(* IEC 61131-3 sources: programs/VI-54/VI-54_20171205/VI-54_20171205/Stations/PLC_VI54/VI-54_171014/Class/_DriveASyncPara, 1 file *)

(* ---- _DriveASyncPara.st ---- *)
#include "..\..\Class\_DriveMngBase\SDDDefinitions.h"

(*!
<Class
	Name               = "_DriveASyncPara"
	Revision           = "1.2"
	RealtimeTask       = "false"
	CyclicTask         = "false"
	BackgroundTask     = "false"
	Sigmatek           = "true"
	OSInterface        = "false"
	HighPriority       = "false"
	Automatic          = "false"
	UpdateMode         = "Prescan"
	IconPath           = ".\Class\_DriveMngBase\Drive.ico"
	SharedCommandTable = "true"
	Objectsize         = "(330,120)"
	Comment            = "class for asynchron parameter handling">
	<Channels>
		<Server Name="ErrorQuit" Visualized="true" Initialize="false" WriteProtected="false" Retentive="false" Comment="quit an error if the asnychron parameter handling failed"/>
		<Server Name="ParaNr" Visualized="true" Initialize="false" WriteProtected="false" Retentive="false" Comment="write the parameter number to read/write the value"/>
		<Server Name="ParaRdWr" Visualized="true" Initialize="false" WriteProtected="false" Retentive="false" Comment="0 .. read the value of the parameter number&#13;&#10;1 .. write a new value of the parameter number"/>
		<Server Name="ParaValue" Visualized="true" Initialize="false" WriteProtected="false" Retentive="false" Comment="Read Command = actual value of the parameter&#13;&#10;Write Command = the new value which has to written to the parameter"/>
		<Server Name="State" Visualized="true" Initialize="false" WriteProtected="true" Retentive="false" Comment="Actual state of the asynchron handling class&#13;&#10;Following states are possible :&#13;&#10;READY&#13;&#10;BUSY&#13;&#10;ERROR"/>
		<Client Name="DriveAxis" Required="true" Internal="false" Comment="object channel to the class _DriveAxis"/>
		<Client Name="ErrorCode" Required="false" Internal="false" Comment="Following error codes are possible :&#13;&#10;ErrorCode &#13;&#10;   3 =    object change only in disable state&#13;&#10;   4 =    object value greater max value or smaller min value&#13;&#10;   5 =    object write not possible&#13;&#10;   6 =    object cannot be changed in this mode&#13;&#10;   7 =    object not available&#13;&#10;   8 =    object read not possible&#13;&#10;   9 =    initialisation processed successful&#13;&#10;  10 =    communication not initialised&#13;&#10;  11 =    axis is not available&#13;&#10;&#13;&#10;"/>
	</Channels>
	<Dependencies>
		<Files>
			<File Path=".\Class\_DriveMngBase\SDDDefinitions.h" Include="true"/>
		</Files>
	</Dependencies>
	<RevDoku>
		<Owner Company="Sigmatek" Author="HasHan"/>
		<Dokumentation Revision="1.2" Date="17.09.2012" Author="RamAnd" Company="Sigmatek" Description="Added method IsOnline to check online state before starting a request."/>
		<Dokumentation Revision="1.1" Date="21.07.2011" Author="RamAnd" Company="Sigmatek" Description="Changed object client DriveAxis from class _DriveAxis to _DriveAxisBase, like in all other drive classes with a connection to the axis object."/>
		<Dokumentation Revision="1.0" Date="05.08.2009" Author="HasHan" Company="Sigmatek" Description="Creation"/>
	</RevDoku>
</Class>
*)
_DriveASyncPara : CLASS
  //Servers:
	State 	: SvrChCmd_iprStates;
	ParaNr 	: SvrCh_DINT;
	ParaRdWr 	: SvrCh_DINT;
	ParaValue 	: SvrCh_DINT;
	ErrorQuit 	: SvrCh_DINT;
  //Clients:
	DriveAxis 	: CltChCmd__DriveAxisBase;
	ErrorCode 	: CltCh_DINT;
  //Variables:
  //Functions:

	FUNCTION VIRTUAL GLOBAL Init;
				//! <Function Comment="get the online state (checks if the axis module can be accessed)" Name="IsOnline"/>
	FUNCTION GLOBAL IsOnline
		VAR_OUTPUT
			OnlineState 	: DINT;			//! <Variable Comment="0..offline&#13;&#10;1..online" Name="IsOnline.OnlineState"/>
		END_VAR;

	FUNCTION VIRTUAL GLOBAL State::NewInst
		VAR_INPUT
			pPara 	: ^CmdStruct;
			pResult 	: ^results;
		END_VAR
		VAR_OUTPUT
			ret_code 	: iprStates;
		END_VAR;

	FUNCTION VIRTUAL GLOBAL ParaNr::Write
		VAR_INPUT
			input (EAX) 	: DINT;
		END_VAR
		VAR_OUTPUT
			result (EAX) 	: DINT;
		END_VAR;

	FUNCTION VIRTUAL GLOBAL ErrorQuit::Write
		VAR_INPUT
			input (EAX) 	: DINT;
		END_VAR
		VAR_OUTPUT
			result (EAX) 	: DINT;
		END_VAR;
  //Tables:
	FUNCTION @STD
		VAR_OUTPUT
			ret_code	: CONFSTATES;
		END_VAR;
	FUNCTION GLOBAL TAB @CT_;
END_CLASS;

#pragma usingLtd _DriveAxisBase

FUNCTION VIRTUAL GLOBAL _DriveASyncPara::Init

	if _firstscan then
    State := READY;
    ErrorCode := 0;
	end_if;

END_FUNCTION

FUNCTION VIRTUAL GLOBAL _DriveASyncPara::State::NewInst
	VAR_INPUT
		pPara 	: ^CmdStruct;
		pResult 	: ^results;
	END_VAR
	VAR_OUTPUT
		ret_code 	: iprStates;
	END_VAR

	ret_code:= READY;

	case pPara^.uiCmd of
	SDD_ASYNC_READY :
		// was the command a read or a write command
		if pPara^.aPara[1] = 0 then
			// read command
			ParaValue := pPara^.aPara[2];
		end_if;
		State := READY;

  SDD_ASYNC_ERROR :
    ErrorCode := pPara^.aPara[1];
    ErrorCode.write(ErrorCode);
    State := ERROR;

	end_case;

END_FUNCTION

FUNCTION VIRTUAL GLOBAL _DriveASyncPara::ParaNr::Write
	VAR_INPUT
		input (EAX) 	: DINT;
	END_VAR
	VAR_OUTPUT
		result (EAX) 	: DINT;
	END_VAR
  VAR
  	IntState    : iprStates;
  END_VAR

	result := ACCESS_DENIED;

	if (State = READY) then
		ParaNr := input;
    IntState := DriveAxis.CmdState.Read();

    if IntState = ERROR then
      if DriveAxis.AxisState.NoHW = 1 then
        ErrorCode := 11;
        ErrorCode.write(ErrorCode);
      end_if;
      State := DriveAxis := IntState;
      return;
    end_if;

		// Add the entry into the ring buffer
		result := DriveAxis.AddASyncEntry(to_usint(ParaNr), to_usint(ParaRdWr), ParaValue, this, 0);
		if result = 0 then
			State := BUSY;
		end_if;
	end_if;

END_FUNCTION

FUNCTION VIRTUAL GLOBAL _DriveASyncPara::ErrorQuit::Write
	VAR_INPUT
		input (EAX) 	: DINT;
	END_VAR
	VAR_OUTPUT
		result (EAX) 	: DINT;
	END_VAR
  VAR
    bError      : BOOL;
    IntState    : iprStates;
  END_VAR

  bError := TRUE;
  // quit an error
  if input = 1 then

    if State = ERROR then
      case ErrorCode of

      11 : //axis is not available
        IntState := DriveAxis.CmdState.Read();
        if IntState = ERROR then
          if DriveAxis.AxisState.NoHW = 0 then
              bError := FALSE;
          end_if;
        end_if;
      else
        bError := FALSE;
      end_case;
    end_if;
  end_if;

  if bError = FALSE then
    State := DriveAxis := READY;
    ErrorCode := 0;
    ErrorCode.write(ErrorCode);
  end_if;

  ErrorQuit := 0;
 	result := ErrorQuit;

END_FUNCTION

FUNCTION GLOBAL _DriveASyncPara::IsOnline
	VAR_OUTPUT
		OnlineState 	: DINT;
	END_VAR

  OnlineState := DriveAxis.Online.Read();

END_FUNCTION
